FUNCTION_BLOCK FB_TankSensors
VAR_IN_OUT
	stTankLevel	:	ST_Tank_Level	;
END_VAR
VAR_INPUT
	volume: REAL:=100; //litr
	//Level
	senHL				:	BOOL	;
	senLL				:	BOOL	;
	nSensorLvl_ID		: 	E_ASense_Name	;
	nSensorLvl_Raw		:	INT		;
	//Temperature
	nSensorTemp_ID		: 	E_ASense_Name	;
	nSensorTemp_Raw		:	INT		;
END_VAR
VAR_OUTPUT
	act_Volume			: REAL;
END_VAR
VAR
	stASensLvl			:	REFERENCE TO ST_AnalogSensor	;
	
	stASensTemp			:	REFERENCE TO ST_AnalogSensor	;
	
	Call_TankLevel			:	FB_AnalogSensor	;
	Call_TankTemp			:	FB_AnalogSensor	;
	tonEmpty: TON;
END_VAR

//Call_TankLevel(nSensorID:=nSensorLvl_ID, nRawSensor:=nSensorLvl_Raw );
//Call_TankTemp(nSensorID:=nSensorTemp_ID, nRawSensor:=nSensorTemp_Raw );
act_TankLvl();
act_Volume:=stTankLevel.rTankLevel;

ACTION act_TankLvl:
stASensLvl REF=g_AnalogSensor.stAnalogSensor[nSensorLvl_ID];

IF stTankLevel.bIn_LL_signal=FALSE AND stTankLevel.bIn_HL_signal=FALSE THEN
	tonEmpty.IN:=TRUE;
ELSE;
	tonEmpty.IN:=FALSE;
END_IF
IF stTankLevel.bIn_LL_signal=TRUE AND stTankLevel.bIn_HL_signal=FALSE THEN
	stTankLevel.e_state:=E_Tank_Level.eLL;
ELSIF stTankLevel.bIn_LL_signal=TRUE AND stTankLevel.bIn_HL_signal=TRUE THEN
	stTankLevel.e_state:=E_Tank_Level.eHL;
ELSIF stTankLevel.bIn_LL_signal=FALSE AND stTankLevel.bIn_HL_signal=TRUE THEN
	stTankLevel.e_state:=E_Tank_Level.eERROR;
END_IF

stTankLevel.rTankLevel:=stASensLvl.Value;
stTankLevel.rTankLevelPercentage:=stTankLevel.rTankLevel/volume*100;
stTankLevel.bIn_HL_signal:=senHL;
stTankLevel.bIn_LL_signal:=senLL;

tonEmpty(PT:=T#3S);
IF tonEmpty.Q THEN;
	stTankLevel.e_state:=E_Tank_Level.eEmpty;
END_IF
END_ACTION

METHOD get_stTankLevel : ST_Tank_Level
VAR_INPUT
END_VAR
VAR
	blank: ST_Tank_Level;
END_VAR
IF __ISVALIDREF(stTankLevel) THEN;
	get_stTankLevel:=stTankLevel;
ELSE;
	get_stTankLevel:=blank;
END_IF
END_METHOD

METHOD get_stTankLevel_OverFlow : BOOL
VAR_INPUT
END_VAR
VAR
	blank: ST_Tank_Level;
END_VAR
IF __ISVALIDREF(stTankLevel) THEN;
	IF stTankLevel.bIn_HL_signal 
	OR stTankLevel.rTankLevelPercentage>100
	OR (NOT MAIN.bTemp_Water_Overweight_check)
	THEN;
		get_stTankLevel_OverFlow:=TRUE;
	ELSE;
		get_stTankLevel_OverFlow:=FALSE;
	END_IF	
ELSE;
	get_stTankLevel_OverFlow:=FALSE;
END_IF
END_METHOD

END_FUNCTION_BLOCK

(* stored: Version 1.1.0.1, ProductVersion 3.1.4024.15
   POU FB_TankSensors: Id {3b995b33-c693-4ceb-8bd6-f0dd6e1df1dc}, SpecialFunc None
   Action act_TankLvl: Id {97fbc1d5-579a-4896-bb72-4b1494685121}
   Method get_stTankLevel: Id {ebb28d4f-5ba4-4bcd-b99d-9ce82e080c07}
   Method get_stTankLevel_OverFlow: Id {577bbcc6-3c21-40bc-aa52-4760d6cb7846} *)
